(* CODESYS project P_Configuration.xml

Project tree, tasks and I/O mapping:
*)

// P_Configuration
PROPERTY P_Configuration : REFERENCE TO ST_AlarmHmiConfiguration
END_PROPERTY
